Fanuc KAREL source: KC00065.KL

PROGRAM KC00065
%NOLOCKGROUP
%ENVIRONMENT CVIS
VAR
  I: INTEGER
  J: INTEGER
  K: INTEGER
  R: REAL
  B: BOOLEAN
  S: STRING[80]
  T: STRING[80]
  P: PATH
  Q: PATH
  AI: ARRAY[8] OF INTEGER
  AB: ARRAY[244] OF BYTE
BEGIN
  V_RALC_QUEUE(I,J,K)
END KC00065
